PROGRAM MBUS_WZaehler_ShopFloor (* hier wird die Klemme, an welche der M-Bus mit den Zählern angeschlossen ist, alle 10ms aufgerufen *)
VAR
	Komm_Klemme_WZaehlerShopFloor	: FB_MBUSKL6781;
	WMZ1xx							: FB_MBUS_General_Ext;
	WMZ2xx							: FB_MBUS_General_Ext;
	WMZ136							: FB_MBUS_General_Ext;
	WMZ236							: FB_MBUS_General_Ext;
	WMZ436							: FB_MBUS_General_Ext;


	adrWMZ1xx			: ST_MBus_SecAdr := (udiIdNumber:=16#50951434); 
	adrWMZ2xx			: ST_MBus_SecAdr := (udiIdNumber:=16#50951428);//DC Schaltschrank
	
	adrWMZ136			: ST_MBus_SecAdr := (udiIdNumber:=16#63350363); //air heat pump CN
	adrWMZ236			: ST_MBus_SecAdr := (udiIdNumber:=16#63350367); //air heat pump HNLT
	adrWMZ436			: ST_MBus_SecAdr := (udiIdNumber:=16#63350353); //air heat pump: heat pump - buffer

END_VAR

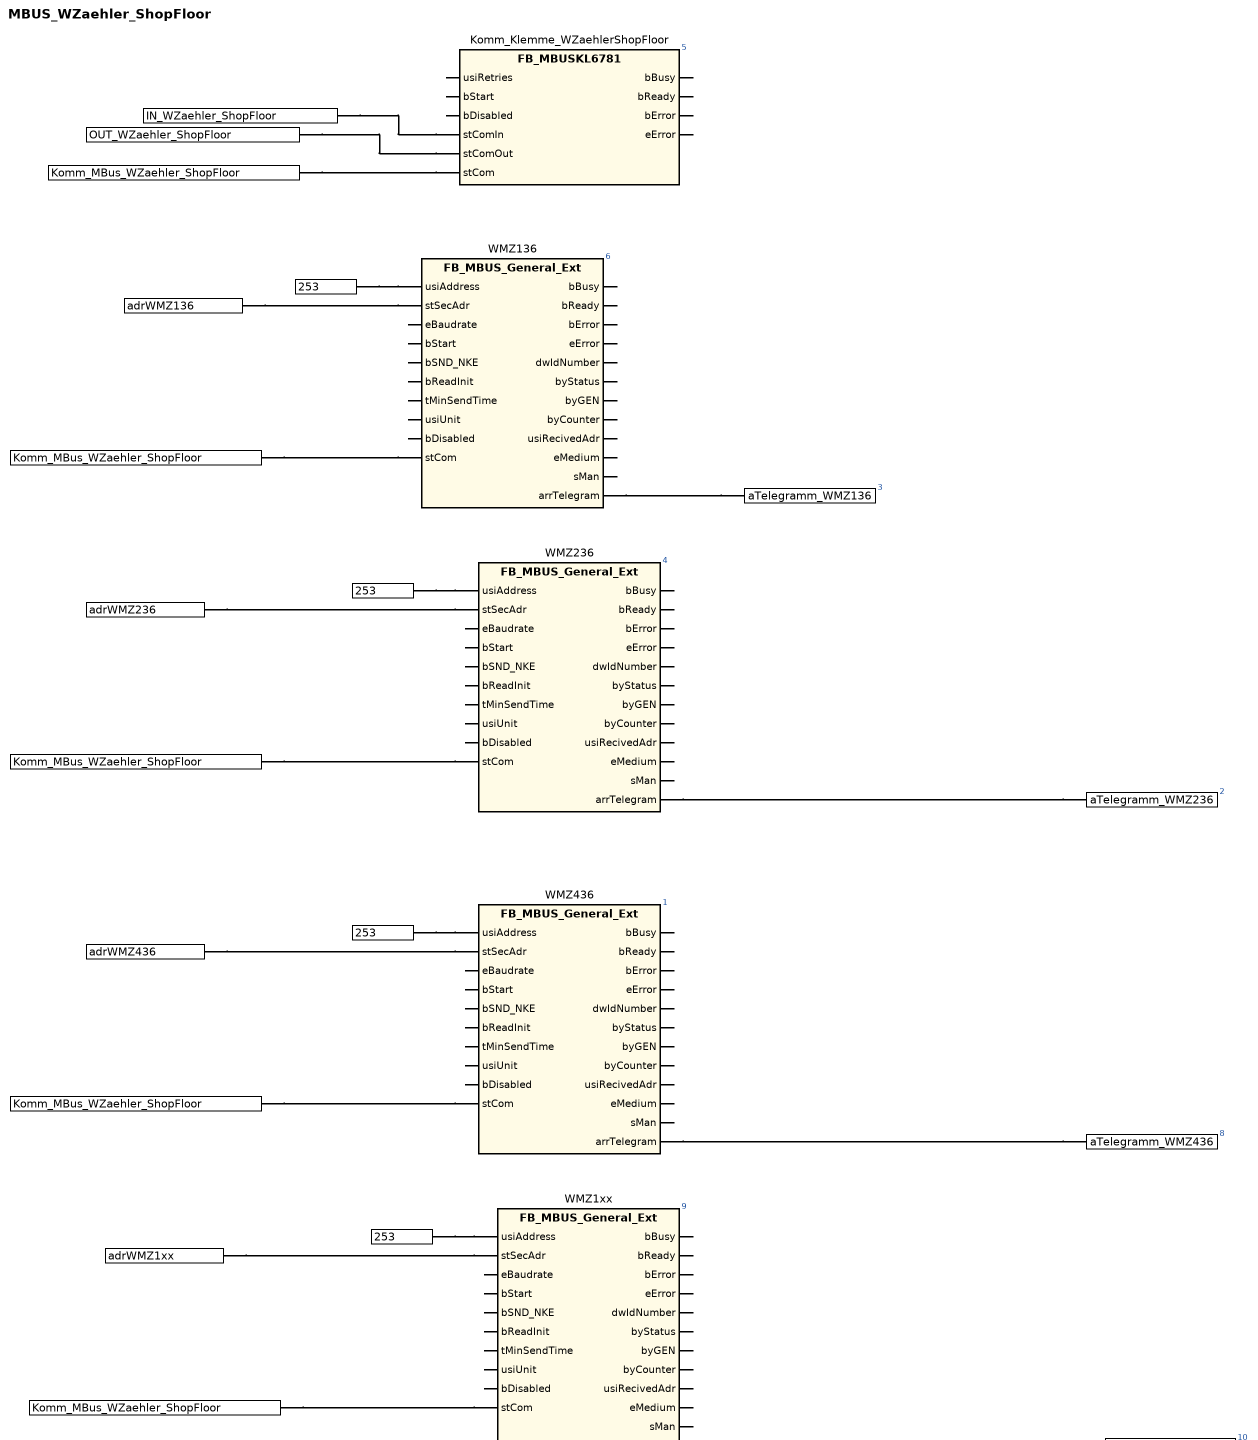
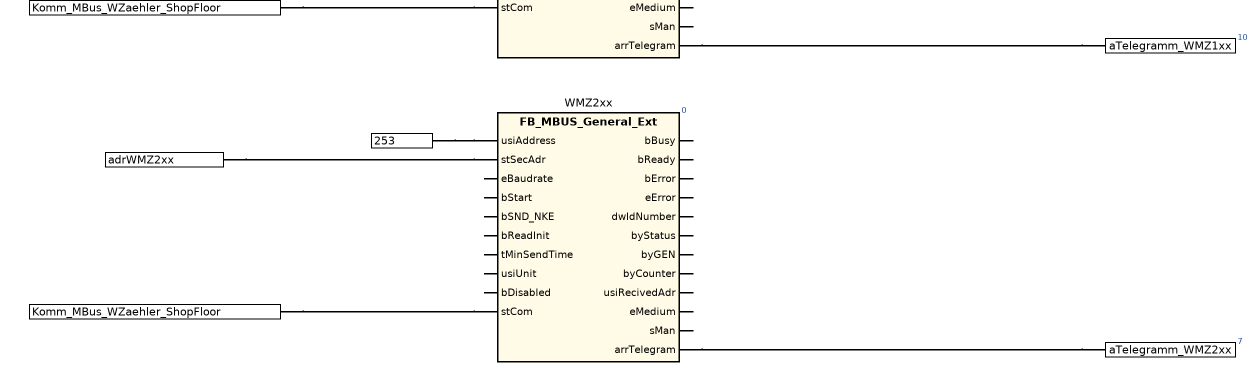
WMZ2xx(usiAddress := 253, stSecAdr := adrWMZ2xx, stCom := Komm_MBus_WZaehler_ShopFloor); // FB_MBUS_General_Ext
WMZ436(usiAddress := 253, stSecAdr := adrWMZ436, stCom := Komm_MBus_WZaehler_ShopFloor); // FB_MBUS_General_Ext
aTelegramm_WMZ236 := WMZ236.arrTelegram;
aTelegramm_WMZ136 := WMZ136.arrTelegram;
WMZ236(usiAddress := 253, stSecAdr := adrWMZ236, stCom := Komm_MBus_WZaehler_ShopFloor); // FB_MBUS_General_Ext
Komm_Klemme_WZaehlerShopFloor(
    stComIn := IN_WZaehler_ShopFloor,
    stComOut := OUT_WZaehler_ShopFloor,
    stCom := Komm_MBus_WZaehler_ShopFloor); // FB_MBUSKL6781
WMZ136(usiAddress := 253, stSecAdr := adrWMZ136, stCom := Komm_MBus_WZaehler_ShopFloor); // FB_MBUS_General_Ext
aTelegramm_WMZ2xx := WMZ2xx.arrTelegram;
aTelegramm_WMZ436 := WMZ436.arrTelegram;
WMZ1xx(usiAddress := 253, stSecAdr := adrWMZ1xx, stCom := Komm_MBus_WZaehler_ShopFloor); // FB_MBUS_General_Ext
aTelegramm_WMZ1xx := WMZ1xx.arrTelegram;

END_PROGRAM

(* stored: Version 1.1.0.1
   POU MBUS_WZaehler_ShopFloor: Id {c5b774f5-c786-4e03-8e02-52a520834700}, SpecialFunc None *)
